Staubli VAL3: new.pgx

public program new(bool& x_bToSave)
  local string l_sNmae
  local bool l_bResult
begin
  l_bResult=userPagePrompt("输入新建名称：",l_sNmae)
  if l_bResult
    if !isDefined(progTemp:pProgItem[l_sNmae])
      insert(progTemp:pProgItem[l_sNmae])
      x_bToSave=true
    endIf
  endIf
end
